Fanuc KAREL source: ka00215.KL

-- PROVISIONAL review KL for V770-1; original PC SHA256 1abe141939d06365f2630a5e77085e96ead051f99a6308161b9ce4472ce5c01e
-- Incomplete behavior may be omitted. Consult companion uncertainty JSON. Do not deploy.
PROGRAM KA00215
%NOLOCKGROUP
BEGIN
  -- UNRESOLVED_PC offsets 5-19; opcodes 22,22,1E
  -- UNRESOLVED_PC offsets 24-28; opcodes 7F
END KA00215
